// Handwritten input matching the prior independent oracle.
TYPE "OracleUnit" VERSION : 0.1 STRUCT ready: BOOL; code: BYTE; count: WORD; END_STRUCT; END_TYPE
DATA_BLOCK "OfficialPadding"
{ S7_Optimized_Access := 'FALSE' }
VAR
a: BYTE; b: BYTE; c: BYTE; bytes: ARRAY[0..6] OF BYTE; tail: BYTE;
END_VAR
BEGIN
END_DATA_BLOCK
DATA_BLOCK "Scalars"
{ S7_Optimized_Access := 'FALSE' }
VAR
b0: BOOL; b1: BOOL; b2: BOOL; b3: BOOL; b4: BOOL; b5: BOOL; b6: BOOL; b7: BOOL; b8: BOOL; octet: BYTE; small: USINT; character: CHAR; signed: INT; unsigned: UINT; bits: WORD; long: DINT; positive: UDINT; mask: DWORD; value: REAL;
END_VAR
BEGIN
END_DATA_BLOCK
DATA_BLOCK "Nested"
{ S7_Optimized_Access := 'FALSE' }
VAR
lead: BYTE; inner: STRUCT a: BOOL; b: BYTE; child: STRUCT u: WORD; flag: BOOL; END_STRUCT; tail: BYTE; END_STRUCT; next: USINT;
END_VAR
BEGIN
END_DATA_BLOCK
DATA_BLOCK "Arrays"
{ S7_Optimized_Access := 'FALSE' }
VAR
lead: BYTE; flags: ARRAY[-2..6] OF BOOL; bytes: ARRAY[3..5] OF BYTE; words: ARRAY[-1..0] OF WORD; values: ARRAY[5..6] OF REAL; items: ARRAY[1..2] OF STRUCT octet: BYTE; flag: BOOL; END_STRUCT; units: ARRAY[-1..0] OF "OracleUnit"; tail: BYTE;
END_VAR
BEGIN
END_DATA_BLOCK
